Fanuc KAREL source: KA00199.KL

PROGRAM KA00199
%NOLOCKGROUP
VAR
  SRC: ARRAY[4] OF VECTOR
  DST: ARRAY[4] OF INTEGER
BEGIN
  DST = SRC
END KA00199
